// TIA Portal V20 export
DATA_BLOCK "OVLADANI_LASER_DB"   // DB400
// stored: AutoNumber false, InstanceOfName OVLADANI_LASER, InstanceOfType FB
"OVLADANI_LASER"
   // VAR
   //    SQCR : Int;
   //    SQCR_WHILE : Int;
   //    SET_WHILE : Bool;
   //    NAZEV_PROGRAMU : String[20];
   //    DELKA_STRINGU : Int;
   //    CHAR_K_ZAPISU : Array[0..71] of Char;
   // END_VAR
BEGIN
END_DATA_BLOCK
